FUNCTION_BLOCK NextFeedHorizonDiag_HMI (* Service Interface Function Block Type *)
  (* Standard: 61499-2 *)
  (* Version 0.0, 10/6/2026, Schneider Electric, template *)
  PACKAGE SE.Nereda;
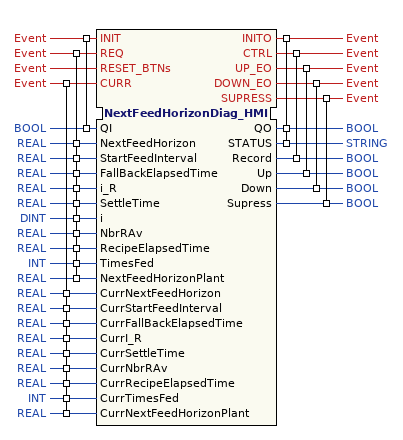
  EVENT_INPUT
    INIT WITH QI;
    REQ WITH NextFeedHorizon, StartFeedInterval, FallBackElapsedTime, i_R, SettleTime, i, NbrRAv, TimesFed, RecipeElapsedTime, NextFeedHorizonPlant;
    RESET_BTNs;
    CURR WITH CurrNextFeedHorizon, CurrStartFeedInterval, CurrFallBackElapsedTime, CurrI_R, CurrSettleTime, CurrNbrRAv, CurrTimesFed, CurrRecipeElapsedTime, CurrNextFeedHorizonPlant;
  END_EVENT
  EVENT_OUTPUT
    INITO WITH QO, STATUS;
    CTRL WITH Record;
    UP_EO WITH Up;
    DOWN_EO WITH Down;
    SUPRESS WITH Supress;
  END_EVENT
  VAR_INPUT
    QI : BOOL;
    NextFeedHorizon : REAL;
    StartFeedInterval : REAL;
    FallBackElapsedTime : REAL;
    i_R : REAL;
    SettleTime : REAL;
    i : DINT;
    NbrRAv : REAL;
    RecipeElapsedTime : REAL;
    TimesFed : INT;
    NextFeedHorizonPlant : REAL;
    CurrNextFeedHorizon : REAL;
    CurrStartFeedInterval : REAL;
    CurrFallBackElapsedTime : REAL;
    CurrI_R : REAL;
    CurrSettleTime : REAL;
    CurrNbrRAv : REAL;
    CurrRecipeElapsedTime : REAL;
    CurrTimesFed : INT;
    CurrNextFeedHorizonPlant : REAL;
  END_VAR
  VAR_OUTPUT
    QO : BOOL; (* Event Output Qualifier *)
    STATUS : STRING; (* Service Status *)
    Record : BOOL;
    Up : BOOL;
    Down : BOOL;
    Supress : BOOL;
  END_VAR
  SERVICE /
    SEQUENCE 
    END_SEQUENCE
  END_SERVICE
END_FUNCTION_BLOCK
